Fanuc KAREL source: kc00035.KL

-- PROVISIONAL review KL for V940-1; original PC SHA256 2c4993aa21cf4dcc8398784f4947464f5ae296f3f84eed4e67d21fcdf5ddc866
-- Incomplete behavior may be omitted. Consult companion uncertainty JSON. Do not deploy.
PROGRAM KC00035
%NOLOCKGROUP
BEGIN
  -- V9_ZERO_TABLE_METADATA_HINT layout=0002_ascii; no indexed target words; source/name/runtime held
  -- UNRESOLVED_PC offsets 5-41; opcodes 27,22,22,2A,22,22,22,31
  -- UNRESOLVED_PC offsets 46-50; opcodes 7F
END KC00035
